Staubli VAL3: main.pgx

program main()
begin
  close(tCurrentTool)
  pPointRx.config.shoulder = lefty
  pPointRx.config.elbow = epositive
  pPointRx.config.wrist = wpositive
  pPointRx2.config.shoulder = lefty
  pPointRx2.config.elbow = epositive
  pPointRx2.config.wrist = wpositive
  mCurrentSpeed.tvel = 100.00
  mCurrentSpeed.blend = joint
  mCurrentSpeed.reach = 0.010
  mCurrentSpeed.leave = 0.010
  call MoveLine(-607.850,543.849,363.215,136.262,30.757,-130.375)
  call MoveJoint(1.00000,-10.00000,20.00000,0.00000,30.00000,0.00000)
  call MoveJoint(2.00000,-10.00000,20.00000,0.00000,30.00000,0.00000)
  call MoveJoint(3.00000,-10.00000,20.00000,0.00000,30.00000,0.00000)

end
